{attribute 'qualified_only'}
VAR_GLOBAL CONSTANT
    stMainLight : ST_LightDefinition := (sLocationCode := 'H-L1-09', sLocationSlug := 'workshop', sLocationName := 'Workshop', sId := 'main', sName := 'Main', nButtonIndex := 1);
END_VAR

(* stored: Version 1.1.0.1
   GVL GVL_WorkshopConfig: Id {c1144eab-69a6-471d-9ccf-4fbd267442a0} *)
